Fanuc KAREL source: ko00059.KL

-- PROVISIONAL review KL for V770-1; original PC SHA256 c7cdff29c8791d4dc97d7a48871634082677ff2e70a6f3a623e9b14f9fe682d5
-- Incomplete behavior may be omitted. Consult companion uncertainty JSON. Do not deploy.
PROGRAM KO00059
%NOLOCKGROUP
BEGIN
  -- UNRESOLVED_PC offsets 5-12; opcodes 9D,23
  -- UNRESOLVED_PC offsets 17-69; opcodes 27,27,49,7E,AD,27,49,7E,AD,22,31,7E,4A
  -- UNRESOLVED_PC offsets 74-78; opcodes 7F
END KO00059
